VAR_GLOBAL
  NULL : PVOID := 0;
END_VAR

(* stored: Version 1.1.0.1
   GVL Constants: Id {eef88d9a-bb0c-4a22-9393-3a929d0f7a35} *)
